(* IEC 61131-3 sources: kns-port-domestic/tools/plcopen/tests/fixtures/constructs/src/DUTs/Motor/Status, 1 file *)

(* ---- ST_MotorSts.dut.st ---- *)
// Состояние двигателя для HMI (DUT во вложенной папке Motor/Status)
TYPE ST_MotorSts :
STRUCT
    xRun : BOOL;
    uiStarts : UINT;
    eMode : E_Mode := E_Mode.OutOfService;
END_STRUCT
END_TYPE
